(* IEC 61131-3 sources: Caravan/Archiv/12-04-19/Stations/MachineControl/MachineControl/Class/InputChange, 1 file *)

(* ---- InputChange.st ---- *)
(*!
<Class
	Name               = "InputChange"
	Revision           = "0.0"
	RealtimeTask       = "false"
	CyclicTask         = "true"
	DefCyclictime      = "100 ms"
	BackgroundTask     = "false"
	Sigmatek           = "false"
	OSInterface        = "false"
	HighPriority       = "false"
	Automatic          = "false"
	UpdateMode         = "Prescan"
	SharedCommandTable = "true"
	Objectsize         = "(284,120)">
	<Channels>
		<Server Name="Out1" Visualized="false" Initialize="false" WriteProtected="false" Retentive="false"/>
		<Server Name="Out2" Visualized="false" Initialize="false" WriteProtected="false" Retentive="false"/>
		<Server Name="Out3" Visualized="false" Initialize="false" WriteProtected="false" Retentive="false"/>
		<Server Name="Out4" Visualized="false" Initialize="false" WriteProtected="false" Retentive="false"/>
		<Client Name="Input1" Required="true" Internal="false"/>
		<Client Name="Input2" Required="true" Internal="false"/>
		<Client Name="Input3" Required="true" Internal="false"/>
		<Client Name="Input4" Required="true" Internal="false"/>
	</Channels>
</Class>
*)
InputChange : CLASS
  //Servers:
	Out1 	: SvrChCmd_DINT;
	Out2 	: SvrCh_DINT;
	Out3 	: SvrCh_DINT;
	Out4 	: SvrCh_DINT;
  //Clients:
	Input1 	: CltCh_DINT;
	Input2 	: CltCh_DINT;
	Input3 	: CltCh_DINT;
	Input4 	: CltCh_DINT;
  //Variables:
  //Functions:

	FUNCTION VIRTUAL GLOBAL CyWork
		VAR_INPUT
			EAX 	: UDINT;
		END_VAR
		VAR_OUTPUT
			state (EAX) 	: UDINT;
		END_VAR;
  //Tables:
	FUNCTION @STD
		VAR_OUTPUT
			ret_code	: CONFSTATES;
		END_VAR;
	FUNCTION GLOBAL TAB @CT_;
END_CLASS;

FUNCTION VIRTUAL GLOBAL InputChange::CyWork
	VAR_INPUT
		EAX 	: UDINT;
	END_VAR
	VAR_OUTPUT
		state (EAX) 	: UDINT;
	END_VAR

  //Read Vars

    Input1  :=  Input1.Read();
    Input2  :=  Input2.Read();
    Input3  :=  Input3.Read();
    Input4  :=  Input4.Read();

    if Input1 = 1 then

        Out1.Write(input:=0);

      else

        out1.Write(input:=1);

    end_if;

    if Input2 = 1 then

        Out2.Write(input:=0);

      else

        out2.Write(input:=1);

    end_if;

    if Input3 = 1 then

        Out3.Write(input:=0);

      else

        out3.Write(input:=1);

    end_if;

    if Input4 = 1 then

        Out4.Write(input:=0);

      else

        out4.Write(input:=1);

    end_if;

	state := READY;

END_FUNCTION
